// Mitsubishi GX Works2 project: DATN_AGV_1   PLC: Q04UDEH

PROGRAM MAIN
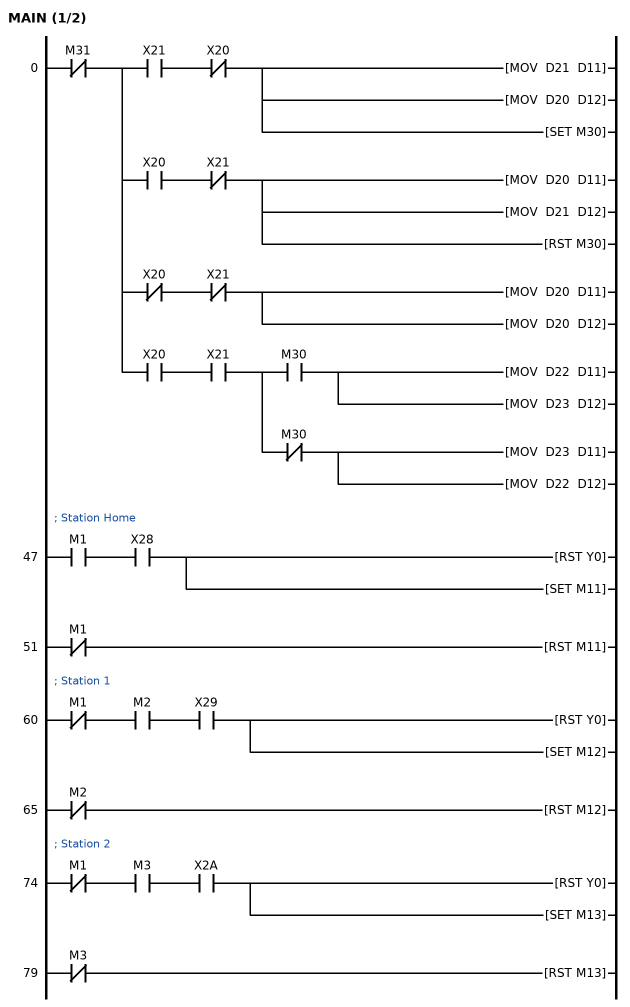
0     LDI     M31
      MPS
      AND     X21
      ANI     X20
      MOV     D21 D11
      MOV     D20 D12
      SET     M30
      MRD
      AND     X20
      ANI     X21
      MOV     D20 D11
      MOV     D21 D12
      RST     M30
      MRD
      ANI     X20
      ANI     X21
      MOV     D20 D11
      MOV     D20 D12
      MPP
      AND     X20
      AND     X21
      MPS
      AND     M30
      MOV     D22 D11
      MOV     D23 D12
      MPP
      ANI     M30
      MOV     D23 D11
      MOV     D22 D12
; Station Home
47    LD      M1
      AND     X28
      RST     Y0
      SET     M11
51    LDI     M1
      RST     M11
; Station 1
60    LDI     M1
      AND     M2
      AND     X29
      RST     Y0
      SET     M12
65    LDI     M2
      RST     M12
; Station 2
74    LDI     M1
      AND     M3
      AND     X2A
      RST     Y0
      SET     M13
79    LDI     M3
      RST     M13
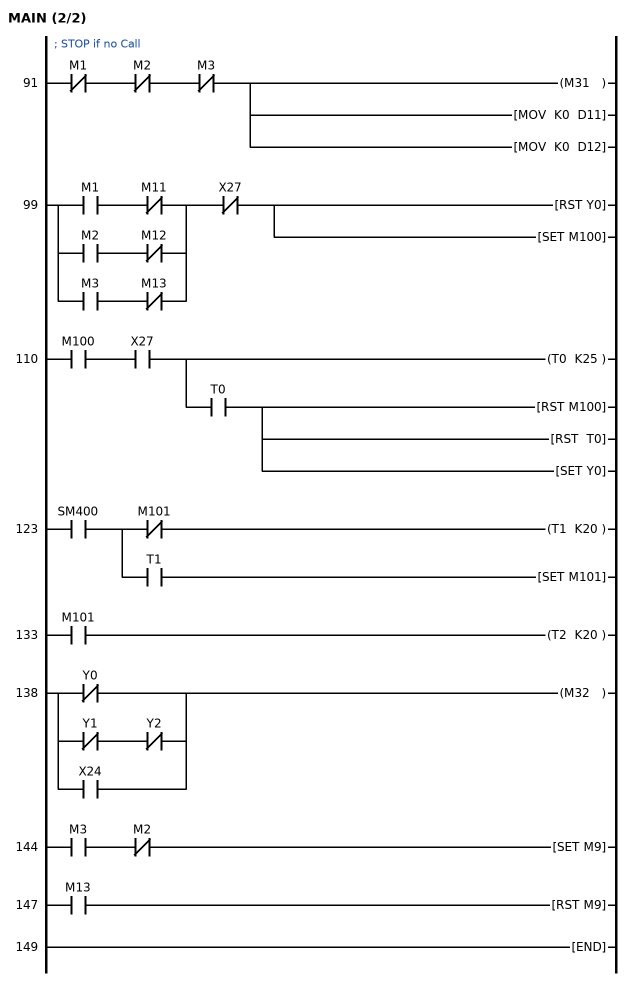
; STOP if no Call
91    LDI     M1
      ANI     M2
      ANI     M3
      OUT     M31
      MOV     K0 D11
      MOV     K0 D12
99    LD      M1
      ANI     M11
      LD      M2
      ANI     M12
      ORB
      LD      M3
      ANI     M13
      ORB
      ANI     X27
      RST     Y0
      SET     M100
110   LD      M100
      AND     X27
      OUT     T0 K25
      AND     T0
      RST     M100
      RST     T0
      SET     Y0
123   LD      SM400
      MPS
      ANI     M101
      OUT     T1 K20
      MPP
      AND     T1
      SET     M101
133   LD      M101
      OUT     T2 K20
138   LDI     Y0
      LDI     Y1
      ANI     Y2
      ORB
      OR      X24
      OUT     M32
144   LD      M3
      ANI     M2
      SET     M9
147   LD      M13
      RST     M9
149   END
END_PROGRAM
